FUNCTION_BLOCK AD2_DWORD_TO_D (* Composite FB for convert DWORD to AD2 *)
  (* Standard: 61499-2; Description: Copyright (c) 2026 HR Agrartechnik GmbH This program and the accompanying materials are made available under the terms of the Eclipse Public License 2.0 which is available at https://www.eclipse.org/legal/epl-2.0/ SPDX-License-Identifier: EPL-2.0 *)
  (* Version 1.0, 2026-11-13, Franz Höpfinger, HR Agrartechnik GmbH, Initial Version - Luecke geschlossen (analog zu AB2_BYTE_TO_B) *)
  PACKAGE adapter::conversion::bidirectional;
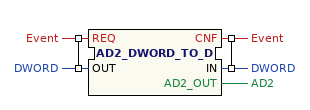
  EVENT_INPUT
    REQ WITH OUT; (* Request to Adapter *)
  END_EVENT
  EVENT_OUTPUT
    CNF WITH IN; (* Confirmation from Adapter *)
  END_EVENT
  VAR_INPUT
    OUT : DWORD; (* Output data to Adapter *)
  END_VAR
  VAR_OUTPUT
    IN : DWORD; (* Input data from Adapter *)
  END_VAR
  PLUGS
    AD2_OUT : adapter::types::bidirectional::AD2; (* Adapter Output *)
  END_PLUGS
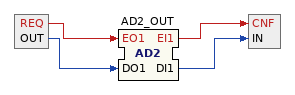
  EVENT_CONNECTIONS
    REQ TO AD2_OUT.EO1;
    AD2_OUT.EI1 TO CNF;
  END_CONNECTIONS
  DATA_CONNECTIONS
    OUT TO AD2_OUT.DO1;
    AD2_OUT.DI1 TO IN;
  END_CONNECTIONS
END_FUNCTION_BLOCK
